ORGANIZATION_BLOCK "Main"
TITLE = Main Program Sweep (Cycle)
{ S7_Optimized_Access := 'TRUE' }
VERSION : 0.1

BEGIN
	"Lampe" := "Taster";
END_ORGANIZATION_BLOCK
